(*
SPDX-FileCopyrightText: c 2026 Oleksandr Tiutyk <trofimich@gmail.com>
SPDX-License-Identifier: MIT
License: https://opensource.org/license/mit
*)

(*!
<summary>Checks independent copies of the configured converter limits.</summary>
<description>
Uses fresh method-local fixtures in a single task cycle.
</description>
*)

{attribute 'no_assign'}
{attribute 'no_explicit_call' := 'do not call this function block directly'}
FUNCTION_BLOCK StaticConverterCopiesLimitsTest EXTENDS TOF_Testing.SingleCycleTest
VAR_STAT
	{attribute 'hide'}
	_ClassName : STRING := __POUNAME();
END_VAR

(*!
<summary>Checks independent copies of the configured converter limits.</summary>
*)
METHOD PROTECTED ExecuteTest
VAR
	minRaw : TOF_Devices_IO.RAW_ANALOG_VALUE;
	maxRaw : TOF_Devices_IO.RAW_ANALOG_VALUE := TOF_Devices_IO.RawAnalogValues.FromInt16(value := 1000);
	converter : TOF_Devices_IO.StaticRangeAnalogValueConverter(
		minAnalogValue := 0.0,
		maxAnalogValue := 100.0,
		minRawValue := minRaw,
		maxRawValue := maxRaw
	);
	resultRaw : TOF_Devices_IO.RAW_ANALOG_VALUE;
END_VAR
// Changing source unions must not change the stored constructor limits.
maxRaw.Int32 := 0;

Assert.ThatLongReal(
	actual := converter.MaxAnalogValue,
	message := "Constructor must preserve the configured analog maximum"
).ToBe(expected := 100.0, tolerance := 0.001);

resultRaw := converter.ConvertAnalogValueToRawValue(
	analogValue := 50.0,
	rawValueType := TOF_Devices_IO.RAW_ANALOG_VALUE_TYPE.INT16
);

Assert.ThatInt(
	actual := resultRaw.Int16,
	message := "Conversion must use copied raw limits after the source changes"
).ToBe(expected := 500);
END_METHOD

//! <summary>Borrows the concrete class name. Callers must not modify it.</summary>
{attribute 'monitoring' := 'call'}
PROPERTY ClassName : REFERENCE TO STRING
GET
ClassName REF= _ClassName;
END_GET
END_PROPERTY

//! <summary>Borrows the compiler-initialized namespace name. Callers must not modify it.</summary>
{attribute 'monitoring' := 'call'}
PROPERTY NamespaceName : REFERENCE TO STRING
GET
NamespaceName REF= CurrentNamespace.Name;
END_GET
END_PROPERTY

//! <summary>Reports the concrete instance size in bytes.</summary>
{attribute 'monitoring' := 'call'}
PROPERTY SelfSize : ULINT
GET
SelfSize := XSIZEOF(THIS^);
END_GET
END_PROPERTY

END_FUNCTION_BLOCK

(* stored: Version 1.1.0.1
   POU StaticConverterCopiesLimitsTest: Id {cc0326de-065d-4c04-9f6b-dc18eeb7e59e}, SpecialFunc None
   Method ExecuteTest: Id {46a68645-e5fa-41bb-8a0b-e2c052a8cd97}
   Property ClassName: Id {fd370106-b7f3-440d-8afe-83cff526ae1b}
   Get Get: Id {352350eb-d115-4bc5-ba19-08779c990264}
   Property NamespaceName: Id {ac059068-bed8-4081-93b1-9172c0c1a0c0}
   Get Get: Id {dc171621-b899-45dd-8702-e1509b4a0473}
   Property SelfSize: Id {cf8499fd-ed0a-4bf7-8a55-a972d07db39f}
   Get Get: Id {7d9c5c8b-693d-4b59-9e9f-6a97ea7c9c3e} *)
